(* IEC 61131-3 sources: genai_codesys/experiments/raw/formal/20261109_234635_2ba96d/public_01/codex_cli__qwen3-coder-flash/attempt_00, 2 files *)

(* ---- declaration.st ---- *)
FUNCTION_BLOCK FB_AutomatedFillingLine
    VAR_INPUT
        bottleSensor : BOOL;
        cleaningConfirmButton : BOOL;
        fillingConfirmButton : BOOL;
        cappingConfirmButton : BOOL;
        packingConfirmButton : BOOL;
        finishedButton : BOOL;
    END_VAR

    VAR_OUTPUT
        Pump_Motor : BOOL;
        Filling_Valve : BOOL;
        Capping_Machine : BOOL;
        Packing_Machine : BOOL;
        Completion_Light : BOOL;
    END_VAR

    VAR
        state : INT := 0;
    END_VAR
END_FUNCTION_BLOCK

(* ---- implementation.st ---- *)
CASE state OF
    0: (* Waiting for bottle *)
        Pump_Motor := bottleSensor;
        IF bottleSensor THEN
            state := 1;
        END_IF;

    1: (* Cleaning *)
        Pump_Motor := TRUE;
        IF cleaningConfirmButton THEN
            state := 2;
        END_IF;

    2: (* Filling *)
        Pump_Motor := FALSE;
        Filling_Valve := TRUE;
        IF fillingConfirmButton THEN
            state := 3;
        END_IF;

    3: (* Capping *)
        Filling_Valve := FALSE;
        Capping_Machine := TRUE;
        IF cappingConfirmButton THEN
            state := 4;
        END_IF;

    4: (* Packaging *)
        Capping_Machine := FALSE;
        Packing_Machine := TRUE;
        IF packingConfirmButton THEN
            state := 5;
        END_IF;

    5: (* Completion *)
        Packing_Machine := FALSE;
        Completion_Light := TRUE;
        IF finishedButton THEN
            state := 0;
        END_IF;

    ELSE
        state := 0;
END_CASE;
